INTERFACE I_DomeState


METHOD CloseCommand : BOOL
END_METHOD


METHOD FoundError : BOOL
END_METHOD


METHOD HomeCommand : BOOL
END_METHOD


METHOD MoveCommand : BOOL
END_METHOD


METHOD OpenCommand : BOOL
END_METHOD


METHOD ParkCommand : BOOL
END_METHOD


METHOD ResetCommand : BOOL
END_METHOD

METHOD RunState : BOOL
VAR_INPUT
END_VAR
END_METHOD


PROPERTY StateID : STRING
GET
END_GET
END_PROPERTY


METHOD StopCommand : BOOL
END_METHOD


METHOD SuccessfulFinished : BOOL
END_METHOD

END_INTERFACE

(* stored: Version 1.1.0.1, ProductVersion 3.1.4024.15
   Itf I_DomeState: Id {b2f6f88a-d56f-445b-bc00-0624b5738555}
   Method CloseCommand: Id {352be468-d16c-467b-8726-c306ee7cd90f}
   Method FoundError: Id {0caae5f8-f18c-4307-9bec-4166c3cd7048}
   Method HomeCommand: Id {4293f3b0-e171-44c9-8fef-6f942c3184b3}
   Method MoveCommand: Id {6e431a8d-905f-42b9-bd77-c182042fe19a}
   Method OpenCommand: Id {1498c54d-e157-48b4-93fc-793d93dafc87}
   Method ParkCommand: Id {1bd7bd84-309d-4e44-9197-c040b737bab3}
   Method ResetCommand: Id {29e0b9ab-e0df-46b5-bed4-b60c365a37ef}
   Method RunState: Id {6706d0a6-a1c6-4fc8-8135-c05165ca8028}
   Property StateID: Id {4d221df5-80db-4dcb-a3c7-2fb94a57b90d}
   Get Get: Id {c4f4c2de-fb35-4b58-88c6-915a0d449a2e}
   Method StopCommand: Id {82ab6c06-0067-49d3-920f-158d61f1c09a}
   Method SuccessfulFinished: Id {ac769bc0-6135-4613-8474-4662273aa323} *)
